FUNCTION_BLOCK FB_House
VAR
    fbLivingRoom : FB_LivingRoom;
    fbLivingRoomCeilingCtrl : FB_LightCtrl;
    fbLivingRoomWallCtrl    : FB_LightCtrl;
    fbLivingRoomAmbientCtrl : FB_LightCtrl;
END_VAR

// Clear all light command inputs before room logic generates commands for this scan.
ClearLightCommands();

// Rooms generate commands for shared devices.
fbLivingRoom();

// Execute all light controllers and light devices once per PLC scan.
ExecuteLights();

METHOD PRIVATE ExecuteLights
// Connect each global light to its relay.
GVL_Lights.fbLivingRoomCeiling(
    stDeviceId := GVL_Lights.stLivingRoomCeilingId,
    iRelay := GVL_Lights.fbLivingRoomCeilingRelay
);
GVL_Lights.fbLivingRoomWall(
    stDeviceId := GVL_Lights.stLivingRoomWallId,
    iRelay := GVL_Lights.fbLivingRoomWallRelay
);
GVL_Lights.fbLivingRoomAmbient(
    stDeviceId := GVL_Lights.stLivingRoomAmbientId,
    iRelay := GVL_Lights.fbLivingRoomAmbientRelay
);

// Execute one controller per light.
fbLivingRoomCeilingCtrl(stLightCmd := GVL_LightCmds.stLivingRoomCeilingCmd, iLight := GVL_Lights.fbLivingRoomCeiling);
fbLivingRoomWallCtrl(stLightCmd := GVL_LightCmds.stLivingRoomWallCmd, iLight := GVL_Lights.fbLivingRoomWall);
fbLivingRoomAmbientCtrl(stLightCmd := GVL_LightCmds.stLivingRoomAmbientCmd, iLight := GVL_Lights.fbLivingRoomAmbient);

// Update relay outputs after command execution in this scan.
GVL_Lights.fbLivingRoomCeilingRelay(stDeviceId := GVL_Lights.stLivingRoomCeilingRelayId);
GVL_Lights.fbLivingRoomWallRelay(stDeviceId := GVL_Lights.stLivingRoomWallRelayId);
GVL_Lights.fbLivingRoomAmbientRelay(stDeviceId := GVL_Lights.stLivingRoomAmbientRelayId);
END_METHOD

METHOD PRIVATE ClearLightCommands
GVL_LightCmds.stLivingRoomCeilingCmd.eAction := E_LightAction.None;
GVL_LightCmds.stLivingRoomCeilingCmd.nBrightness := 0;

GVL_LightCmds.stLivingRoomWallCmd.eAction := E_LightAction.None;
GVL_LightCmds.stLivingRoomWallCmd.nBrightness := 0;

GVL_LightCmds.stLivingRoomAmbientCmd.eAction := E_LightAction.None;
GVL_LightCmds.stLivingRoomAmbientCmd.nBrightness := 0;
END_METHOD

END_FUNCTION_BLOCK

(* stored: Version 1.1.0.1, ProductVersion 3.1.4026.20
   POU FB_House: Id {A8100001-3B71-4C96-8F25-7A1B2C3D4001}
   Method ExecuteLights: Id {A8100001-3B71-4C96-8F25-7A1B2C3D4002}
   Method ClearLightCommands: Id {A8100001-3B71-4C96-8F25-7A1B2C3D4003} *)
